(* IEC 61131-3 sources: trust-platform/manual-tests/clean-root/src, 5 files *)

(* ---- ICounter.st ---- *)
INTERFACE ICounter
    METHOD Next : DINT
    END_METHOD
    PROPERTY Value : DINT
        GET
        END_GET
    END_PROPERTY
END_INTERFACE

(* ---- AddTwo.st ---- *)
FUNCTION AddTwo : DINT
VAR_INPUT
    EN : BOOL := TRUE;
    A : DINT;
    B : DINT;
END_VAR
VAR_OUTPUT
    ENO : BOOL;
END_VAR
IF EN THEN
    ENO := TRUE;
    AddTwo := A + B;
ELSE
    ENO := FALSE;
    AddTwo := DINT#0;
END_IF
END_FUNCTION

(* ---- CounterFb.st ---- *)
FUNCTION_BLOCK CounterFb IMPLEMENTS ICounter
VAR
    x : DINT;
END_VAR

METHOD PUBLIC Next : DINT
    x := x + 1;
    Next := x;
END_METHOD

PUBLIC PROPERTY Value : DINT
    GET
        Value := x;
    END_GET
END_PROPERTY
END_FUNCTION_BLOCK

(* ---- Configuration.st ---- *)
CONFIGURATION CleanConfig
RESOURCE Res1 ON PLC
    TASK FastTask(INTERVAL := T#100ms, PRIORITY := 1);
    PROGRAM P1 WITH FastTask : Main;
END_RESOURCE
END_CONFIGURATION

(* ---- Main2.st ---- *)
PROGRAM Main2
VAR
    counter : CounterFb;
    outVal : DINT;
    ok : BOOL;
END_VAR
outVal := AddTwo(A := 1, B := 2);
outVal := AddTwo(EN := TRUE, A := 1, B := 2, ENO => ok);
outVal := counter.Next();
outVal := counter.Value;
END_PROGRAM
